(* PLC project MotorStarter, plcforge plcforge examples 0.4.0 *)
(* stored: creationDateTime 2026-02-11T09:15:00 *)

FUNCTION_BLOCK MotorStarter
  VAR_INPUT
    startButton : BOOL;  (* Momentary start push button *)
    stopButton : BOOL;  (* Normally closed stop push button *)
    overload : BOOL;  (* Thermal overload contact *)
  END_VAR
  VAR_OUTPUT
    motor : BOOL;  (* Motor contactor *)
    warmedUp : BOOL;  (* Set once the motor has run for the warm-up time *)
  END_VAR
  VAR
    warmUpTimer : TON;
  END_VAR

(* LD diagram, written out as Structured Text *)
motor := (startButton OR motor) AND NOT stopButton AND NOT overload;
warmUpTimer(IN := motor, PT := T#5s);
warmedUp := warmUpTimer.Q;
END_FUNCTION_BLOCK
